(* IEC 61131-3 sources: codesys-to-astra/src/POUs/F_C2aRealToStringFormat, 2 files *)

(* ---- F_C2aRealToStringFormat.decl.st ---- *)
// Назначение: замена OSU.REAL_TO_STRING_FORMAT (OwenStringUtils v3.0, с. 9): REAL -> строка с заданным
//             числом знаков после разделителя (точка или запятая; недопустимый разделитель — точка).
//             |значение| > 1e8 — экспоненциальная запись REAL_TO_STRING. Округление последнего знака может
//             отличаться от ОВЕН (обёртка, исход check).
// Автор:      kr0nsch
// Версия:     0.1.0
// Документ:   docs/LIBMAP.md
FUNCTION F_C2aRealToStringFormat : STRING(80)
VAR_INPUT
    rValueToConvert : REAL;                     // значение
    usiSignificantDigitsCount : USINT;          // знаков после разделителя (0..7)
    eDecimalSeparator : E_C2aDecimalSeparator;  // разделитель
END_VAR
VAR
    usiDigits : USINT;      // знаков после разделителя после ограничения
    lrAbs : LREAL;          // модуль значения
    lrScaled : LREAL;       // модуль · 10^usiDigits + 0.5
    uliPow : ULINT;          // 10 ^ usiDigits
    uliScaled : ULINT;       // модуль, умноженный на 10 ^ usiDigits и округлённый
    uliInt : ULINT;          // целая часть
    uliFrac : ULINT;         // дробная часть
    sFrac : STRING(80);     // дробная часть строкой
    sSep : STRING(1);       // разделитель
    usiIdx : USINT;         // счётчик
END_VAR

(* ---- F_C2aRealToStringFormat.impl.st ---- *)
IF eDecimalSeparator = E_C2aDecimalSeparator.COMMA THEN
    sSep := ',';
ELSE
    sSep := '.';
END_IF
IF ABS(rValueToConvert) > GVL_C2aConst.EXP_THRESHOLD THEN
    F_C2aRealToStringFormat := REAL_TO_STRING(rValueToConvert);
    IF sSep = ',' AND FIND(F_C2aRealToStringFormat, '.') > 0 THEN
        F_C2aRealToStringFormat := REPLACE(F_C2aRealToStringFormat, ',', 1, FIND(F_C2aRealToStringFormat, '.'));
    END_IF
    RETURN;
END_IF
usiDigits := MIN(usiSignificantDigitsCount, GVL_C2aConst.MAX_FRACTION_DIGITS);
uliPow := 1;
FOR usiIdx := 1 TO usiDigits DO
    uliPow := uliPow * 10;  // lint:allow STL008 десятичная система
END_FOR
lrAbs := ABS(REAL_TO_LREAL(rValueToConvert));
lrScaled := lrAbs * ULINT_TO_LREAL(uliPow) + 0.5;  // lint:allow STL008 округление половины вверх
// LREAL_TO_ULINT округляет к ближайшему — приводим к floor(x + 0.5)
uliScaled := LREAL_TO_ULINT(lrScaled);
IF ULINT_TO_LREAL(uliScaled) > lrScaled THEN
    uliScaled := uliScaled - 1;
END_IF
uliInt := uliScaled / uliPow;
uliFrac := uliScaled MOD uliPow;
F_C2aRealToStringFormat := ULINT_TO_STRING(uliInt);
IF usiDigits > 0 THEN
    sFrac := ULINT_TO_STRING(uliFrac);
    WHILE LEN(sFrac) < USINT_TO_INT(usiDigits) DO
        sFrac := CONCAT('0', sFrac);
    END_WHILE
    F_C2aRealToStringFormat := CONCAT(CONCAT(F_C2aRealToStringFormat, sSep), sFrac);
END_IF
IF rValueToConvert < 0.0 AND uliScaled > 0 THEN
    F_C2aRealToStringFormat := CONCAT('-', F_C2aRealToStringFormat);
END_IF
